FUNCTION "LAUER KEYS 2" : VOID
TITLE =Lauer Keys 2
NAME : ZEITEN1
VERSION : 0.0

BEGIN
NETWORK
TITLE =

      OPN   "DB LAUER";

NETWORK
TITLE =

      A     "M 171.0";
      BEC   ;
NETWORK
TITLE =

      AN    "M 151.7";
      JC    M001;
      L     2#100000000;
      T     DBW   72;
M001: NOP   0;
NETWORK
TITLE =

      AN    "M 151.7";
      JC    M002;
      L     2#1001;
      T     DBW   76;
M002: NOP   0;
NETWORK
TITLE =

      A     "M 171.0";
      BEC   ;
NETWORK
TITLE =

      A(    ;
      L     DBB   32;
      L     1;
      ==I   ;
      )     ;
      A     "M 151.7";
      JC    M003;
      JU    M003;

M003: CALL "LAUER TIME" (
           QUEL                     := DBW  240,
           _TIME                    := MW   130);


END_FUNCTION
